PROGRAM Signals
VAR
	fbTimer1: TON;
	fbTimer2: TON;
	fbBlinker: FB_Blinker;	
END_VAR

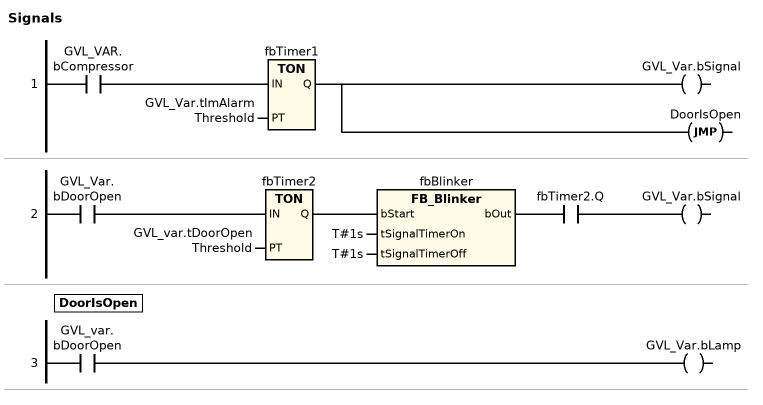
// NETWORK 1
fbTimer1(IN := GVL_VAR.bCompressor, PT := GVL_Var.tImAlarmThreshold); // TON
GVL_Var.bSignal := fbTimer1.Q;
IF fbTimer1.Q THEN JMP DoorIsOpen; END_IF

// NETWORK 2
fbTimer2(IN := GVL_Var.bDoorOpen, PT := GVL_var.tDoorOpenThreshold); // TON
fbBlinker(bStart := fbTimer2.Q, tSignalTimerOn := T#1s, tSignalTimerOff := T#1s); // FB_Blinker
GVL_Var.bSignal := fbBlinker.bOut AND fbTimer2.Q;

// NETWORK 3
DoorIsOpen:
GVL_Var.bLamp := GVL_var.bDoorOpen;

END_PROGRAM

(* stored: Version 1.1.0.1, ProductVersion 3.1.4024.16
   POU Signals: Id {ac6ac33d-86a4-4eff-a91e-1e31d05993f0}, SpecialFunc None *)
